Fanuc KAREL source: KB00062.KL

PROGRAM KB00062
%NOLOCKGROUP
%ENVIRONMENT PBQMGR
VAR
  P1: INTEGER
  P2: QUEUE_TYPE
  P3: ARRAY[4] OF INTEGER
  P4: INTEGER
BEGIN
  P1 = 1
  P3[1] = 1
  P4 = 1
  DELETE_QUEUE(P1, P2, P3, P4)
END KB00062
